Fanuc KAREL source: KD00025.KL

PROGRAM KD00025
%NOLOCKGROUP
VAR
  I: INTEGER
  J: INTEGER
  B: BOOLEAN
  R: REAL
  S: STRING[80]
BEGIN
  CONDITION[1]: WITH $PRIORITY = 50
  WHEN DIN[1] = ON DO
    I = 1
  ENDCONDITION
END KD00025
